(* Logix 5000 project; controller SigmaAldrich vendor 1 type 14 code 77 rev 15.4; software revision 15.02 *)

TASK MainTask (continuous, watchdog 500 ms) : MainProgram

MODULES
   Controller : vendor 1 type 14 code 77 (CompactLogixL32EController 0, rev 15.4)
      LocalENB : 1769-L32E Ethernet Port (CompactLogixL32Ethernet 1, rev 15.3)
      Local : CompactBus (CompactVirtualAdapter 3, rev 15.3, Input RPI 2 ms)
          : vendor 1 type 7 code 69 (Compact 12, rev 3.1, Input RPI 2 ms)
          : vendor 1 type 7 code 69 (Compact 9, rev 3.1, Input RPI 2 ms)
          : vendor 1 type 7 code 69 (Compact 7, rev 3.1, Input RPI 2 ms)
          : vendor 1 type 7 code 69 (Compact 10, rev 3.1, Input RPI 2 ms)
          : vendor 1 type 7 code 69 (Compact 11, rev 3.1, Input RPI 2 ms)
          : vendor 1 type 7 code 69 (Compact 8, rev 3.1, Input RPI 2 ms)
          : 1769-OW16 (Compact 1, rev 1.1, Output RPI 2 ms)
          : 1769-OW16 (Compact 6, rev 1.1, Output RPI 2 ms)
          : 1769-OW16 (Compact 3, rev 1.1, Output RPI 2 ms)
          : 1769-OW16 (Compact 4, rev 1.1, Output RPI 2 ms)
          : 1769-OW16 (Compact 2, rev 1.1, Output RPI 2 ms)
          : 1769-OW16 (Compact 5, rev 1.1, Output RPI 2 ms)
END_MODULES

VAR_GLOBAL   (* controller tags *)
   Airlock_N1002_03_04_E_Stop_OSR : BOOL;
   Airlock_N1002_03_04_Violation_MDI_Bit : BOOL := 1;
   Airlock_N1002_03_04_Violation_MDI_OSR : BOOL := 1;
   Airlock_N1005_E_Stop_OSR : BOOL;
   Airlock_N1005_Violation_MDI_Bit : BOOL;
   Airlock_N1005_Violation_MDI_OSR : BOOL;
   Airlock_N1006_E_Stop_OSR : BOOL;
   Airlock_N1006_Violation_MDI_Bit : BOOL;
   Airlock_N1006_Violation_MDI_OSR : BOOL;
   Airlock_N1008_E_Stop_OSR : BOOL;
   Airlock_N1008_Violation_MDI_Bit : BOOL;
   Airlock_N1008_Violation_MDI_OSR : BOOL;
   Airlock_N1009_E_Stop_OSR : BOOL;
   Airlock_N1009_Violation_MDI_Bit : BOOL;
   Airlock_N1009_Violation_MDI_OSR : BOOL;
   Airlock_N1011_E_Stop_OSR : BOOL;
   Airlock_N1011_Violation_MDI_Bit : BOOL := 1;
   Airlock_N1011_Violation_MDI_OSR : BOOL := 1;
   Airlock_N1012_E_Stop_OSR : BOOL;
   Airlock_N1012_Violation_MDI_Bit : BOOL := 1;
   Airlock_N1012_Violation_MDI_OSR : BOOL := 1;
   Airlock_N1021_E_Stop_OSR : BOOL;
   Airlock_N1021_Violation_MDI_Bit : BOOL;
   Airlock_N1021_Violation_MDI_OSR : BOOL;
   Airlock_N1043_E_Stop_OSR : BOOL;
   Airlock_N1043_Violation_MDI_Bit : BOOL := 1;
   Airlock_N1043_Violation_MDI_OSR : BOOL := 1;
   Airlock_N1044_E_Stop_OSR : BOOL;
   Airlock_N1044_Violation_MDI_Bit : BOOL;
   Airlock_N1044_Violation_MDI_OSR : BOOL;
   Airlock_N1051_54_55_E_Stop_OSR : BOOL;
   Airlock_N1051_54_55_Violation_MDI_Bit : BOOL := 1;
   Airlock_N1051_54_55_Violation_MDI_OSR : BOOL;
   Airlock_N1052_E_Stop_OSR : BOOL;
   Airlock_N1052_Violation_MDI_Bit : BOOL;
   Airlock_N1052_Violation_MDI_OSR : BOOL;
   Airlock_N1065_E_Stop_OSR : BOOL;
   Airlock_N1065_Violation_MDI_Bit : BOOL;
   Airlock_N1065_Violation_MDI_OSR : BOOL;
   Airlock_N1066_E_Stop_OSR : BOOL;
   Airlock_N1066_Violation_MDI_Bit : BOOL := 1;
   Airlock_N1066_Violation_MDI_OSR : BOOL := 1;
   Airlock_N1068_E_Stop_OSR : BOOL;
   Airlock_N1068_Violation_MDI_Bit : BOOL;
   Airlock_N1068_Violation_MDI_OSR : BOOL;
   Annuciator_Bit_Airlock_N1002_03_04 : BOOL := 1;
   Annuciator_Bit_Airlock_N1005 : BOOL;
   Annuciator_Bit_Airlock_N1006 : BOOL;
   Annuciator_Bit_Airlock_N1008 : BOOL;
   Annuciator_Bit_Airlock_N1009 : BOOL;
   Annuciator_Bit_Airlock_N1011 : BOOL := 1;
   Annuciator_Bit_Airlock_N1012 : BOOL := 1;
   Annuciator_Bit_Airlock_N1021 : BOOL;
   Annuciator_Bit_Airlock_N1043 : BOOL := 1;
   Annuciator_Bit_Airlock_N1044 : BOOL;
   Annuciator_Bit_Airlock_N1051_54_55 : BOOL := 1;
   Annuciator_Bit_Airlock_N1052 : BOOL;
   Annuciator_Bit_Airlock_N1065 : BOOL;
   Annuciator_Bit_Airlock_N1066 : BOOL := 1;
   Annuciator_Bit_Airlock_N1068 : BOOL;
   Door_N1002A_Timer : TIMER := (PRE := 30000);
   Door_N1002B_Timer : TIMER := (PRE := 30000);
   Door_N1002C_Timer : TIMER := (PRE := 30000);
   Door_N1003A_Timer : TIMER := (PRE := 30000);
   Door_N1003C_Timer : TIMER := (PRE := 30000, ACC := 30000, EN := 1, DN := 1);
   Door_N1004A_Timer : TIMER := (PRE := 30000);
   Door_N1004B_Timer : TIMER := (PRE := 30000);
   Door_N1005A_Timer : TIMER := (PRE := 30000);
   Door_N1005B_Timer : TIMER := (PRE := 30000);
   Door_N1006A_Timer : TIMER := (PRE := 30000);
   Door_N1006B_Timer : TIMER := (PRE := 30000);
   Door_N1008A_Timer : TIMER := (PRE := 30000);
   Door_N1008B_Timer : TIMER := (PRE := 30000);
   Door_N1009A_Timer : TIMER := (PRE := 30000);
   Door_N1009B_Timer : TIMER := (PRE := 30000);
   Door_N1011A_Timer : TIMER := (PRE := 30000, ACC := 30000, EN := 1, DN := 1);
   Door_N1011B_Timer : TIMER := (PRE := 30000, ACC := 30000, EN := 1, DN := 1);
   Door_N1012_Timer : TIMER := (PRE := 30000, ACC := 30000, EN := 1, DN := 1);
   Door_N1021A_Timer : TIMER := (PRE := 30000);
   Door_N1021B_Timer : TIMER := (PRE := 30000);
   Door_N1021C_Timer : TIMER := (PRE := 30000);
   Door_N1043A_Timer : TIMER := (PRE := 30000, ACC := 30000, EN := 1, DN := 1);
   Door_N1043B_Timer : TIMER := (PRE := 30000);
   Door_N1044A_Timer : TIMER := (PRE := 30000);
   Door_N1044B_Timer : TIMER := (PRE := 30000);
   Door_N1044C_Timer : TIMER := (PRE := 30000);
   Door_N1051A_Timer : TIMER := (PRE := 30000, ACC := 30000, EN := 1, DN := 1);
   Door_N1051B_Timer : TIMER := (PRE := 30000, ACC := 30000, EN := 1, DN := 1);
   Door_N1052A_Timer : TIMER := (PRE := 30000);
   Door_N1052B_Timer : TIMER := (PRE := 30000);
   Door_N1053_Timer : TIMER := (PRE := 30000, ACC := 30000, EN := 1, DN := 1);
   Door_N1054A_Timer : TIMER := (PRE := 30000, ACC := 30000, EN := 1, DN := 1);
   Door_N1054B_Timer : TIMER := (PRE := 30000, ACC := 30000, EN := 1, DN := 1);
   Door_N1054C_Timer : TIMER := (PRE := 30000, ACC := 30000, EN := 1, DN := 1);
   Door_N1055_Timer : TIMER := (PRE := 30000, ACC := 30000, EN := 1, DN := 1);
   Door_N1058B_Timer : TIMER := (PRE := 30000);
   Door_N1065A_Timer : TIMER := (PRE := 30000);
   Door_N1065B_Timer : TIMER := (PRE := 30000);
   Door_N1066A_Timer : TIMER := (PRE := 30000, ACC := 30000, EN := 1, DN := 1);
   Door_N1066B_Timer : TIMER := (PRE := 30000, ACC := 30000, EN := 1, DN := 1);
   Door_N1068A_Timer : TIMER := (PRE := 30000);
   Door_N1068B_Timer : TIMER := (PRE := 30000);
   MDI_Violation_N1002_03_04_Bit : BOOL := 1;
   MDI_Violation_N1005_Bit : BOOL;
   MDI_Violation_N1006_Bit : BOOL;
   MDI_Violation_N1008_Bit : BOOL;
   MDI_Violation_N1009_Bit : BOOL;
   MDI_Violation_N1011_Bit : BOOL := 1;
   MDI_Violation_N1012_Bit : BOOL := 1;
   MDI_Violation_N1021_Bit : BOOL;
   MDI_Violation_N1043_Bit : BOOL := 1;
   MDI_Violation_N1044_Bit : BOOL;
   MDI_Violation_N1051_54_55_Bit : BOOL := 1;
   MDI_Violation_N1052_Bit : BOOL;
   MDI_Violation_N1065_Bit : BOOL;
   MDI_Violation_N1066_Bit : BOOL := 1;
   MDI_Violation_N1068_Bit : BOOL;
   N1002_03_04_Airlock_Latch : BOOL := 1;
   N1002_03_04_Emergency_Release_Latch : BOOL := 1;
   N1005_Airlock_Latch : BOOL;
   N1005_Emergency_Release_Latch : BOOL;
   N1006_Airlock_Latch : BOOL;
   N1006_Emergency_Release_Latch : BOOL;
   N1008_Airlock_Latch : BOOL;
   N1008_Emergency_Release_Latch : BOOL;
   N1009_Airlock_Latch : BOOL;
   N1009_Emergency_Release_Latch : BOOL;
   N1011_Airlock_Latch : BOOL := 1;
   N1011_Emergency_Release_Latch : BOOL;
   N1012_Airlock_Latch : BOOL := 1;
   N1012_Emergency_Release_Latch : BOOL;
   N1021_Airlock_Latch : BOOL;
   N1021_Emergency_Release_Latch : BOOL;
   N1021C_Door_Latch_Bit : BOOL;
   N1043_Airlock_Latch : BOOL;
   N1043_Emergency_Release_Latch : BOOL;
   N1044_Airlock_Latch : BOOL;
   N1044_Emergency_Release_Latch : BOOL;
   N1044A_Door_Latch_Bit : BOOL;
   N1051_54_55_Airlock_Latch : BOOL := 1;
   N1051_54_55_Emergency_Release_Latch : BOOL;
   N1052_Airlock_Latch : BOOL;
   N1052_Emergency_Release_Latch : BOOL;
   N1052A_Door_Latch_Bit : BOOL;
   N1065_Airlock_Latch : BOOL;
   N1065_Emergency_Release_Latch : BOOL;
   N1066_Airlock_Latch : BOOL := 1;
   N1066_Emergency_Release_Latch : BOOL;
   N1068_Airlock_Latch : BOOL;
   N1068_Emergency_Release_Latch : BOOL;
   N1068B_Door_Latch_Bit : BOOL;
END_VAR

PROGRAM MainProgram   (* main routine MainRoutine *)
VAR
   Airlock_N1009_Delay_Tmr : TIMER := (PRE := 2000);
   Airlock_N1009_MDI_Delay_Tmr : TIMER := (PRE := 2000, ACC := 2001, EN := 1, DN := 1);
END_VAR

ROUTINE DI01_N1051_N1054_N0155   (* ladder *)
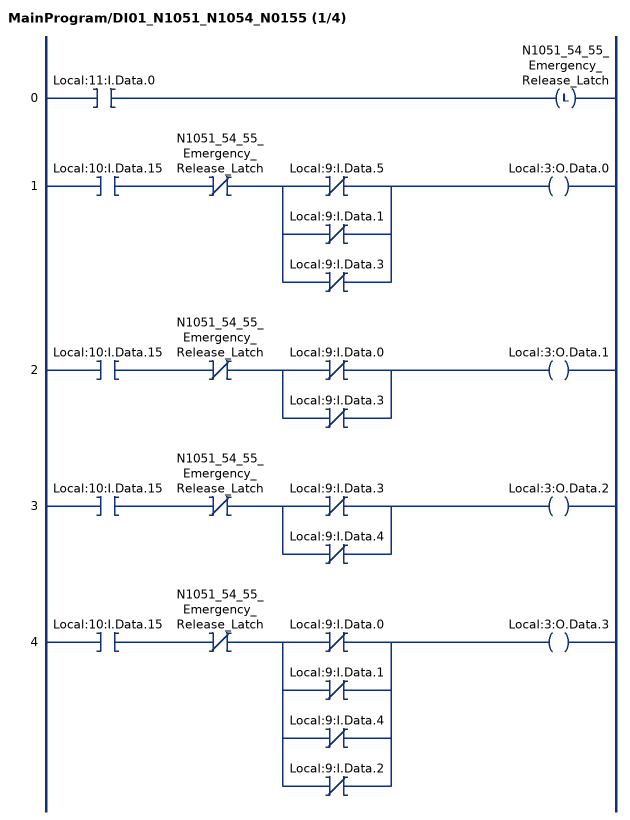
   0: XIC(Local:11:I.Data.0)OTL(N1051_54_55_Emergency_Release_Latch);
   1: XIC(Local:10:I.Data.15)XIO(N1051_54_55_Emergency_Release_Latch)[XIO(Local:9:I.Data.5) ,XIO(Local:9:I.Data.1) ,XIO(Local:9:I.Data.3) ]OTE(Local:3:O.Data.0);
   2: XIC(Local:10:I.Data.15)XIO(N1051_54_55_Emergency_Release_Latch)[XIO(Local:9:I.Data.0) ,XIO(Local:9:I.Data.3) ]OTE(Local:3:O.Data.1);
   3: XIC(Local:10:I.Data.15)XIO(N1051_54_55_Emergency_Release_Latch)[XIO(Local:9:I.Data.3) ,XIO(Local:9:I.Data.4) ]OTE(Local:3:O.Data.2);
   4: XIC(Local:10:I.Data.15)XIO(N1051_54_55_Emergency_Release_Latch)[XIO(Local:9:I.Data.0) ,XIO(Local:9:I.Data.1) ,XIO(Local:9:I.Data.4) ,XIO(Local:9:I.Data.2) ]OTE(Local:3:O.Data.3);
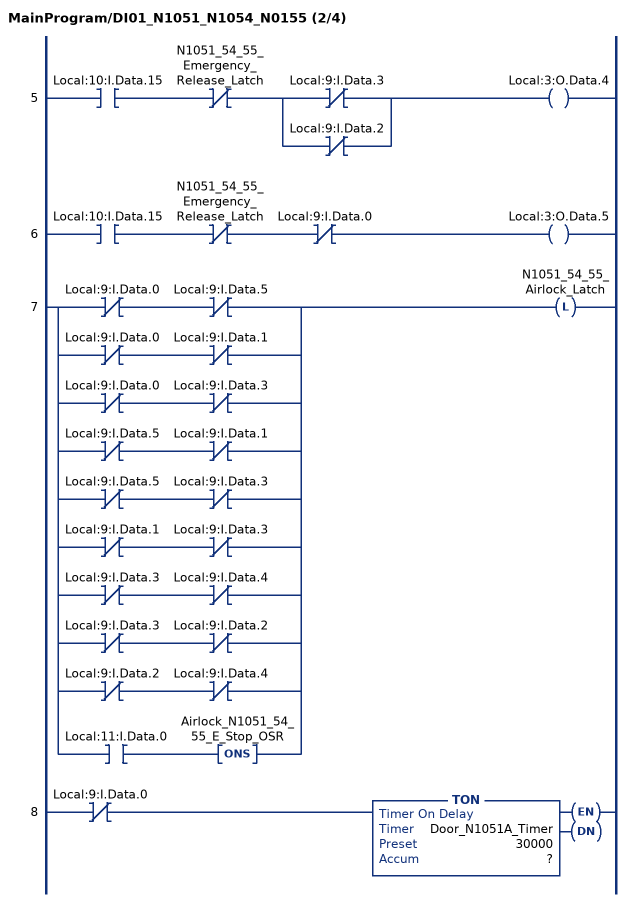
   5: XIC(Local:10:I.Data.15)XIO(N1051_54_55_Emergency_Release_Latch)[XIO(Local:9:I.Data.3) ,XIO(Local:9:I.Data.2) ]OTE(Local:3:O.Data.4);
   6: XIC(Local:10:I.Data.15)XIO(N1051_54_55_Emergency_Release_Latch)XIO(Local:9:I.Data.0)OTE(Local:3:O.Data.5);
   7: [XIO(Local:9:I.Data.0) XIO(Local:9:I.Data.5) ,XIO(Local:9:I.Data.0) XIO(Local:9:I.Data.1) ,XIO(Local:9:I.Data.0) XIO(Local:9:I.Data.3) ,XIO(Local:9:I.Data.5) XIO(Local:9:I.Data.1) ,XIO(Local:9:I.Data.5) XIO(Local:9:I.Data.3) ,XIO(Local:9:I.Data.1) XIO(Local:9:I.Data.3) ,XIO(Local:9:I.Data.3) XIO(Local:9:I.Data.4) ,XIO(Local:9:I.Data.3) XIO(Local:9:I.Data.2) ,XIO(Local:9:I.Data.2) XIO(Local:9:I.Data.4) ,XIC(Local:11:I.Data.0) ONS(Airlock_N1051_54_55_E_Stop_OSR) ]OTL(N1051_54_55_Airlock_Latch);
   8: XIO(Local:9:I.Data.0)TON(Door_N1051A_Timer,?,?);
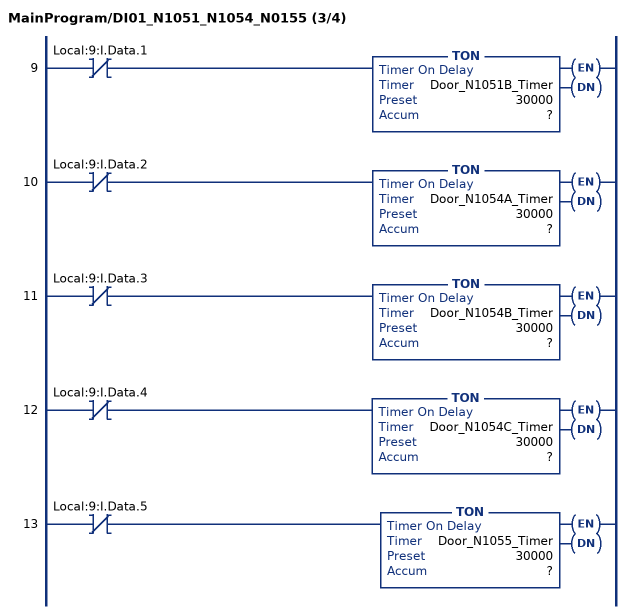
   9: XIO(Local:9:I.Data.1)TON(Door_N1051B_Timer,?,?);
   10: XIO(Local:9:I.Data.2)TON(Door_N1054A_Timer,?,?);
   11: XIO(Local:9:I.Data.3)TON(Door_N1054B_Timer,?,?);
   12: XIO(Local:9:I.Data.4)TON(Door_N1054C_Timer,?,?);
   13: XIO(Local:9:I.Data.5)TON(Door_N1055_Timer,?,?);
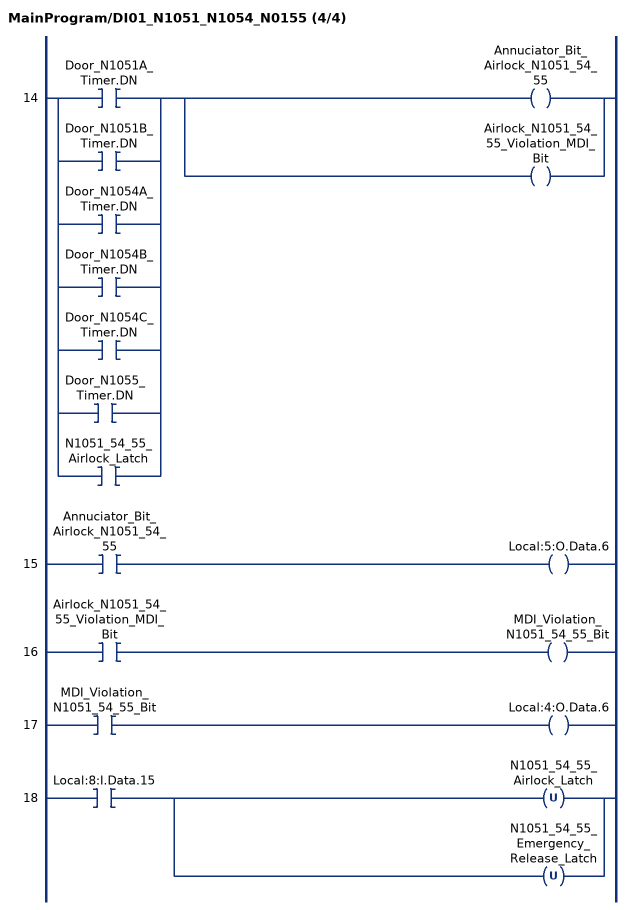
   14: [XIC(Door_N1051A_Timer.DN) ,XIC(Door_N1051B_Timer.DN) ,XIC(Door_N1054A_Timer.DN) ,XIC(Door_N1054B_Timer.DN) ,XIC(Door_N1054C_Timer.DN) ,XIC(Door_N1055_Timer.DN) ,XIC(N1051_54_55_Airlock_Latch) ][OTE(Annuciator_Bit_Airlock_N1051_54_55) ,OTE(Airlock_N1051_54_55_Violation_MDI_Bit) ];
   15: XIC(Annuciator_Bit_Airlock_N1051_54_55)OTE(Local:5:O.Data.6);
   16: XIC(Airlock_N1051_54_55_Violation_MDI_Bit)OTE(MDI_Violation_N1051_54_55_Bit);
   17: XIC(MDI_Violation_N1051_54_55_Bit)OTE(Local:4:O.Data.6);
   18: XIC(Local:8:I.Data.15)[OTU(N1051_54_55_Airlock_Latch) ,OTU(N1051_54_55_Emergency_Release_Latch) ];
END_ROUTINE

ROUTINE DI02_N1002_N1003_N1004   (* ladder *)
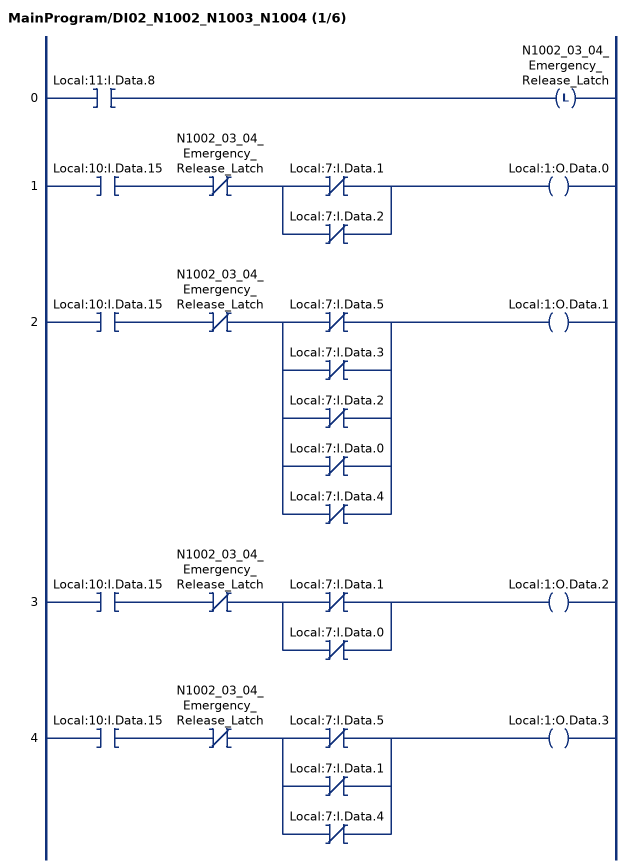
   0: XIC(Local:11:I.Data.8)OTL(N1002_03_04_Emergency_Release_Latch);
   1: XIC(Local:10:I.Data.15)XIO(N1002_03_04_Emergency_Release_Latch)[XIO(Local:7:I.Data.1) ,XIO(Local:7:I.Data.2) ]OTE(Local:1:O.Data.0);
   2: XIC(Local:10:I.Data.15)XIO(N1002_03_04_Emergency_Release_Latch)[XIO(Local:7:I.Data.5) ,XIO(Local:7:I.Data.3) ,XIO(Local:7:I.Data.2) ,XIO(Local:7:I.Data.0) ,XIO(Local:7:I.Data.4) ]OTE(Local:1:O.Data.1);
   3: XIC(Local:10:I.Data.15)XIO(N1002_03_04_Emergency_Release_Latch)[XIO(Local:7:I.Data.1) ,XIO(Local:7:I.Data.0) ]OTE(Local:1:O.Data.2);
   4: XIC(Local:10:I.Data.15)XIO(N1002_03_04_Emergency_Release_Latch)[XIO(Local:7:I.Data.5) ,XIO(Local:7:I.Data.1) ,XIO(Local:7:I.Data.4) ]OTE(Local:1:O.Data.3);
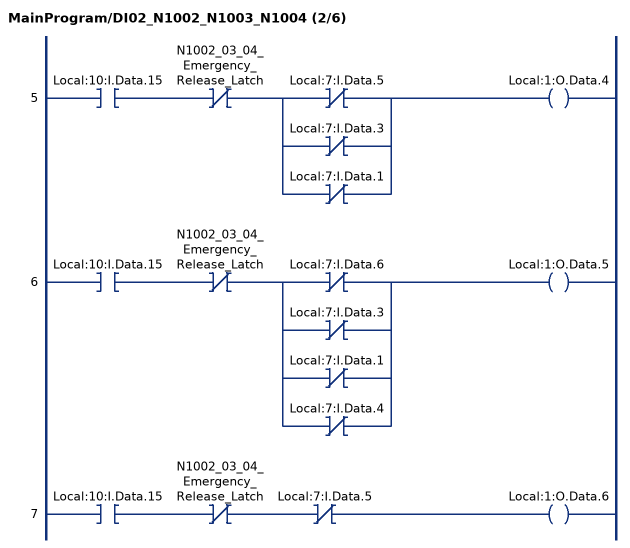
   5: XIC(Local:10:I.Data.15)XIO(N1002_03_04_Emergency_Release_Latch)[XIO(Local:7:I.Data.5) ,XIO(Local:7:I.Data.3) ,XIO(Local:7:I.Data.1) ]OTE(Local:1:O.Data.4);
   6: XIC(Local:10:I.Data.15)XIO(N1002_03_04_Emergency_Release_Latch)[XIO(Local:7:I.Data.6) ,XIO(Local:7:I.Data.3) ,XIO(Local:7:I.Data.1) ,XIO(Local:7:I.Data.4) ]OTE(Local:1:O.Data.5);
   7: XIC(Local:10:I.Data.15)XIO(N1002_03_04_Emergency_Release_Latch)XIO(Local:7:I.Data.5)OTE(Local:1:O.Data.6);
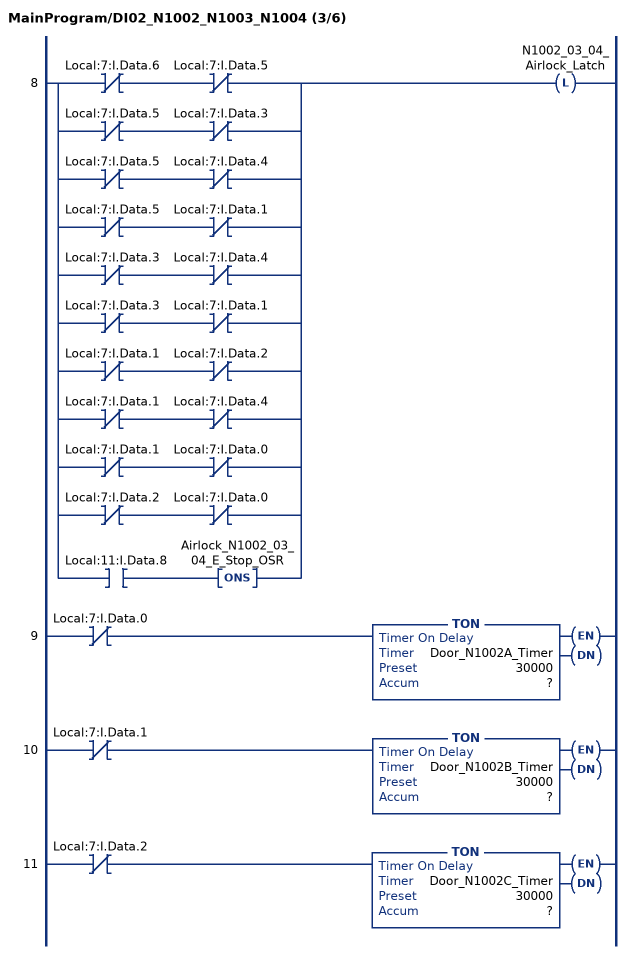
   8: [XIO(Local:7:I.Data.6) XIO(Local:7:I.Data.5) ,XIO(Local:7:I.Data.5) XIO(Local:7:I.Data.3) ,XIO(Local:7:I.Data.5) XIO(Local:7:I.Data.4) ,XIO(Local:7:I.Data.5) XIO(Local:7:I.Data.1) ,XIO(Local:7:I.Data.3) XIO(Local:7:I.Data.4) ,XIO(Local:7:I.Data.3) XIO(Local:7:I.Data.1) ,XIO(Local:7:I.Data.1) XIO(Local:7:I.Data.2) ,XIO(Local:7:I.Data.1) XIO(Local:7:I.Data.4) ,XIO(Local:7:I.Data.1) XIO(Local:7:I.Data.0) ,XIO(Local:7:I.Data.2) XIO(Local:7:I.Data.0) ,XIC(Local:11:I.Data.8) ONS(Airlock_N1002_03_04_E_Stop_OSR) ]OTL(N1002_03_04_Airlock_Latch);
   9: XIO(Local:7:I.Data.0)TON(Door_N1002A_Timer,?,?);
   10: XIO(Local:7:I.Data.1)TON(Door_N1002B_Timer,?,?);
   11: XIO(Local:7:I.Data.2)TON(Door_N1002C_Timer,?,?);
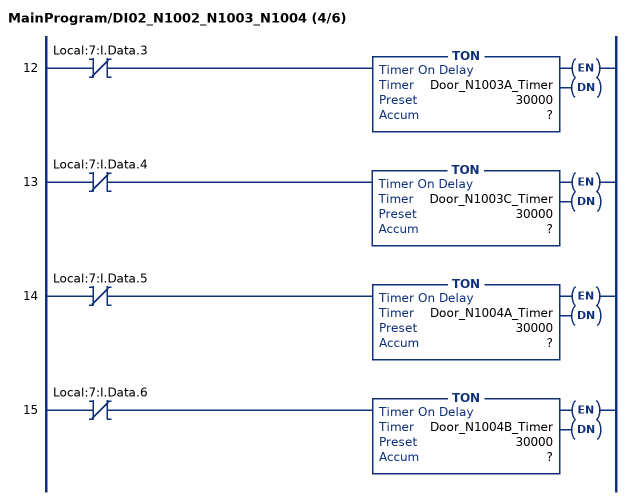
   12: XIO(Local:7:I.Data.3)TON(Door_N1003A_Timer,?,?);
   13: XIO(Local:7:I.Data.4)TON(Door_N1003C_Timer,?,?);
   14: XIO(Local:7:I.Data.5)TON(Door_N1004A_Timer,?,?);
   15: XIO(Local:7:I.Data.6)TON(Door_N1004B_Timer,?,?);
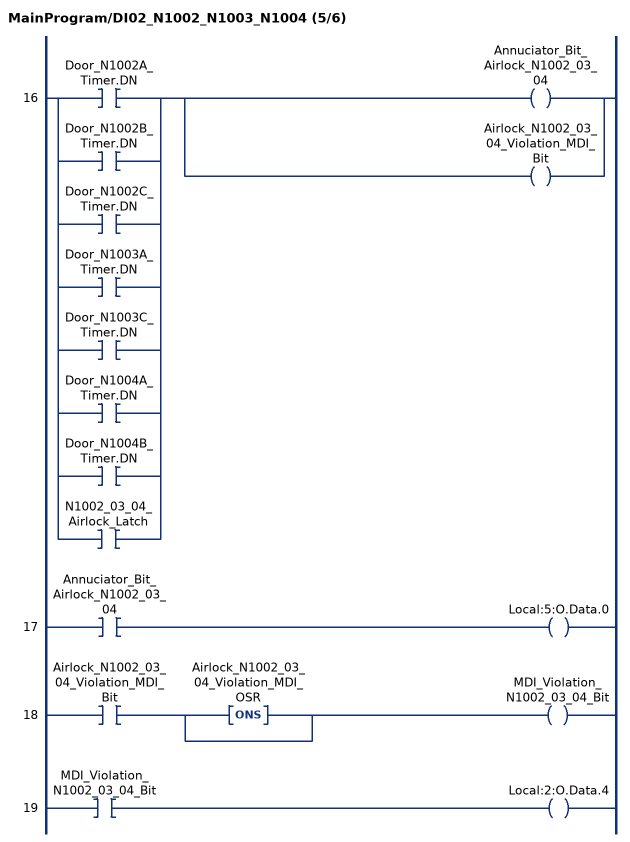
   16: [XIC(Door_N1002A_Timer.DN) ,XIC(Door_N1002B_Timer.DN) ,XIC(Door_N1002C_Timer.DN) ,XIC(Door_N1003A_Timer.DN) ,XIC(Door_N1003C_Timer.DN) ,XIC(Door_N1004A_Timer.DN) ,XIC(Door_N1004B_Timer.DN) ,XIC(N1002_03_04_Airlock_Latch) ][OTE(Annuciator_Bit_Airlock_N1002_03_04) ,OTE(Airlock_N1002_03_04_Violation_MDI_Bit) ];
   17: XIC(Annuciator_Bit_Airlock_N1002_03_04)OTE(Local:5:O.Data.0);
   18: XIC(Airlock_N1002_03_04_Violation_MDI_Bit)[ONS(Airlock_N1002_03_04_Violation_MDI_OSR) ,]OTE(MDI_Violation_N1002_03_04_Bit);
   19: XIC(MDI_Violation_N1002_03_04_Bit)OTE(Local:2:O.Data.4);
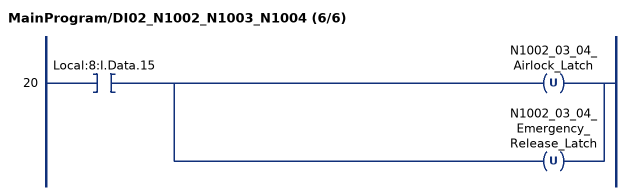
   20: XIC(Local:8:I.Data.15)[OTU(N1002_03_04_Airlock_Latch) ,OTU(N1002_03_04_Emergency_Release_Latch) ];
END_ROUTINE

ROUTINE DI03_N1021   (* ladder *)
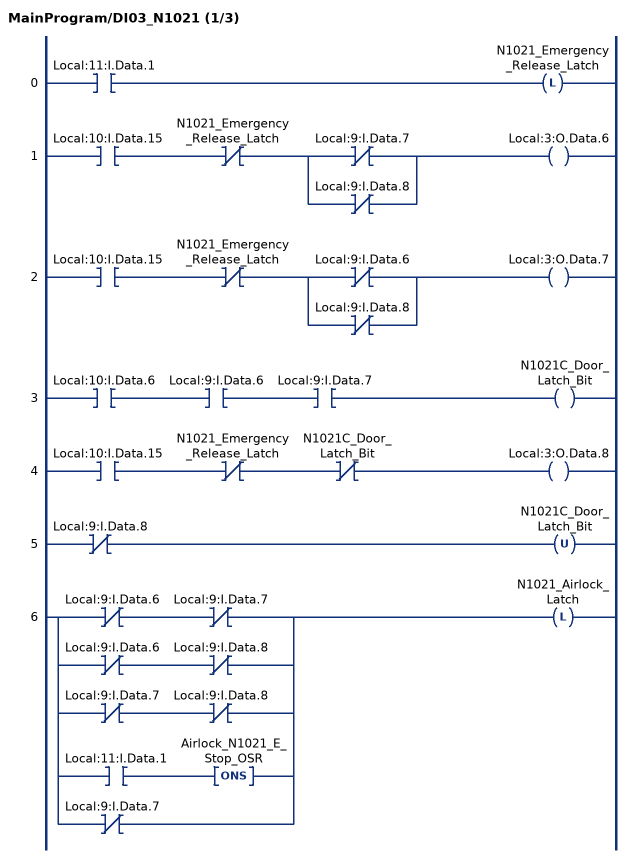
   0: XIC(Local:11:I.Data.1)OTL(N1021_Emergency_Release_Latch);
   1: XIC(Local:10:I.Data.15)XIO(N1021_Emergency_Release_Latch)[XIO(Local:9:I.Data.7) ,XIO(Local:9:I.Data.8) ]OTE(Local:3:O.Data.6);
   2: XIC(Local:10:I.Data.15)XIO(N1021_Emergency_Release_Latch)[XIO(Local:9:I.Data.6) ,XIO(Local:9:I.Data.8) ]OTE(Local:3:O.Data.7);
   3: XIC(Local:10:I.Data.6)XIC(Local:9:I.Data.6)XIC(Local:9:I.Data.7)OTE(N1021C_Door_Latch_Bit);
   4: XIC(Local:10:I.Data.15)XIO(N1021_Emergency_Release_Latch)XIO(N1021C_Door_Latch_Bit)OTE(Local:3:O.Data.8);
   5: XIO(Local:9:I.Data.8)OTU(N1021C_Door_Latch_Bit);
   6: [XIO(Local:9:I.Data.6) XIO(Local:9:I.Data.7) ,XIO(Local:9:I.Data.6) XIO(Local:9:I.Data.8) ,XIO(Local:9:I.Data.7) XIO(Local:9:I.Data.8) ,XIC(Local:11:I.Data.1) ONS(Airlock_N1021_E_Stop_OSR) ,XIO(Local:9:I.Data.7) ]OTL(N1021_Airlock_Latch);
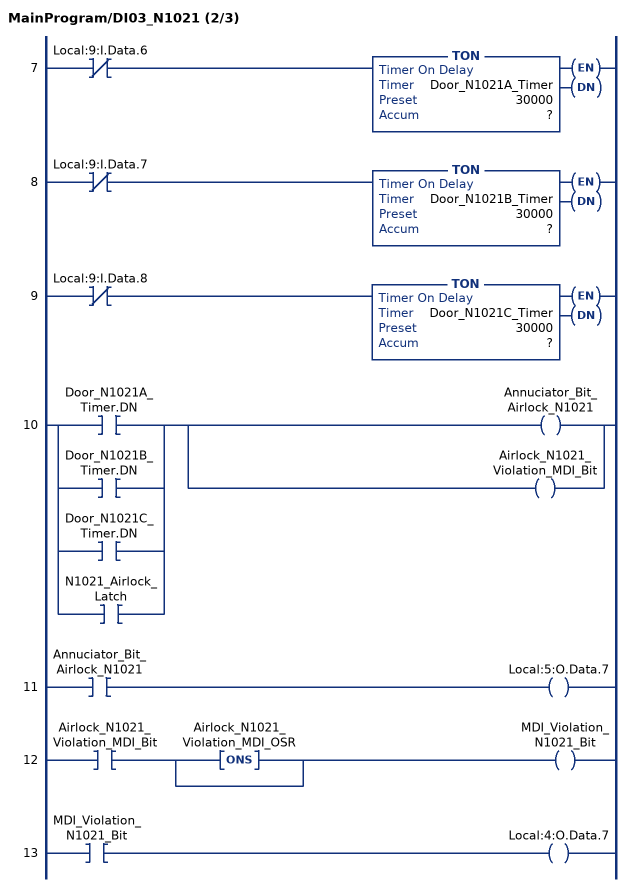
   7: XIO(Local:9:I.Data.6)TON(Door_N1021A_Timer,?,?);
   8: XIO(Local:9:I.Data.7)TON(Door_N1021B_Timer,?,?);
   9: XIO(Local:9:I.Data.8)TON(Door_N1021C_Timer,?,?);
   10: [XIC(Door_N1021A_Timer.DN) ,XIC(Door_N1021B_Timer.DN) ,XIC(Door_N1021C_Timer.DN) ,XIC(N1021_Airlock_Latch) ][OTE(Annuciator_Bit_Airlock_N1021) ,OTE(Airlock_N1021_Violation_MDI_Bit) ];
   11: XIC(Annuciator_Bit_Airlock_N1021)OTE(Local:5:O.Data.7);
   12: XIC(Airlock_N1021_Violation_MDI_Bit)[ONS(Airlock_N1021_Violation_MDI_OSR) ,]OTE(MDI_Violation_N1021_Bit);
   13: XIC(MDI_Violation_N1021_Bit)OTE(Local:4:O.Data.7);
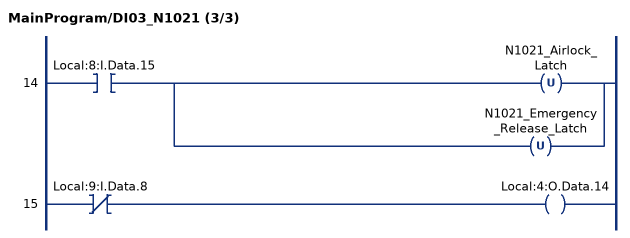
   14: XIC(Local:8:I.Data.15)[OTU(N1021_Airlock_Latch) ,OTU(N1021_Emergency_Release_Latch) ];
   15: XIO(Local:9:I.Data.8)OTE(Local:4:O.Data.14);
END_ROUTINE

ROUTINE DI04_N1005   (* ladder *)
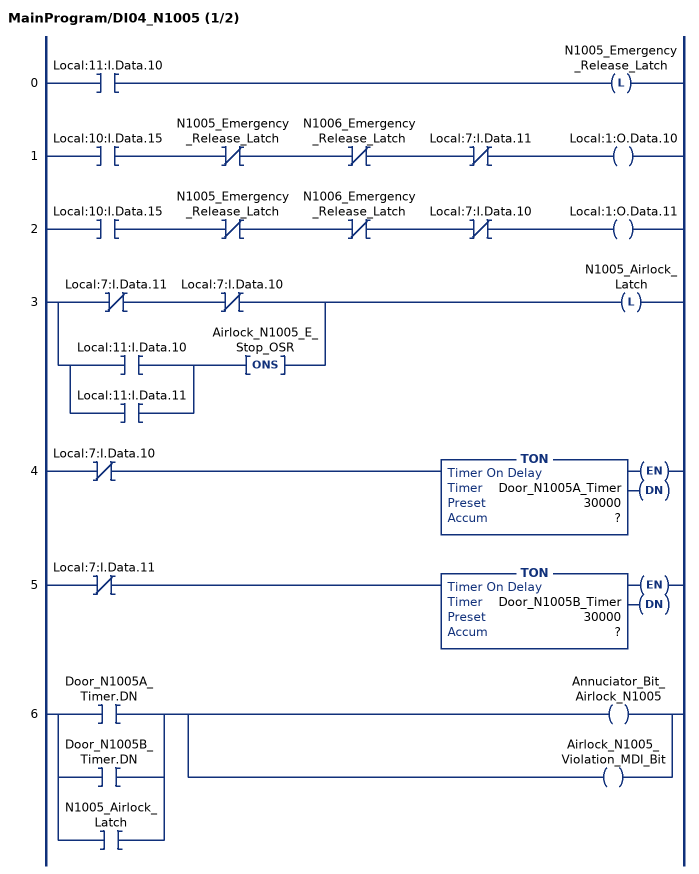
   0: XIC(Local:11:I.Data.10)OTL(N1005_Emergency_Release_Latch);
   1: XIC(Local:10:I.Data.15)XIO(N1005_Emergency_Release_Latch)XIO(N1006_Emergency_Release_Latch)XIO(Local:7:I.Data.11)OTE(Local:1:O.Data.10);
   2: XIC(Local:10:I.Data.15)XIO(N1005_Emergency_Release_Latch)XIO(N1006_Emergency_Release_Latch)XIO(Local:7:I.Data.10)OTE(Local:1:O.Data.11);
   3: [XIO(Local:7:I.Data.11) XIO(Local:7:I.Data.10) ,[XIC(Local:11:I.Data.10) ,XIC(Local:11:I.Data.11) ] ONS(Airlock_N1005_E_Stop_OSR) ]OTL(N1005_Airlock_Latch);
   4: XIO(Local:7:I.Data.10)TON(Door_N1005A_Timer,?,?);
   5: XIO(Local:7:I.Data.11)TON(Door_N1005B_Timer,?,?);
   6: [XIC(Door_N1005A_Timer.DN) ,XIC(Door_N1005B_Timer.DN) ,XIC(N1005_Airlock_Latch) ][OTE(Annuciator_Bit_Airlock_N1005) ,OTE(Airlock_N1005_Violation_MDI_Bit) ];
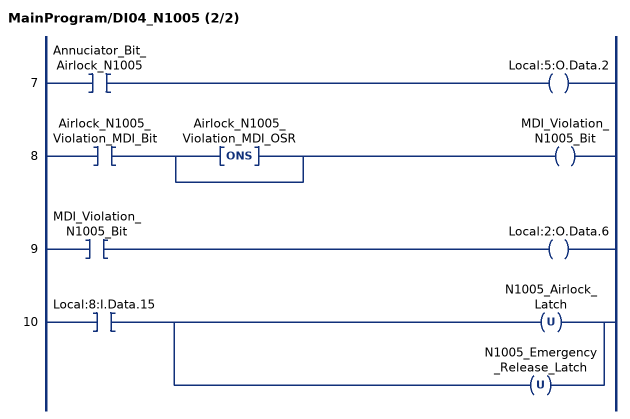
   7: XIC(Annuciator_Bit_Airlock_N1005)OTE(Local:5:O.Data.2);
   8: XIC(Airlock_N1005_Violation_MDI_Bit)[ONS(Airlock_N1005_Violation_MDI_OSR) ,]OTE(MDI_Violation_N1005_Bit);
   9: XIC(MDI_Violation_N1005_Bit)OTE(Local:2:O.Data.6);
   10: XIC(Local:8:I.Data.15)[OTU(N1005_Airlock_Latch) ,OTU(N1005_Emergency_Release_Latch) ];
END_ROUTINE

ROUTINE DI05_N1006   (* ladder *)
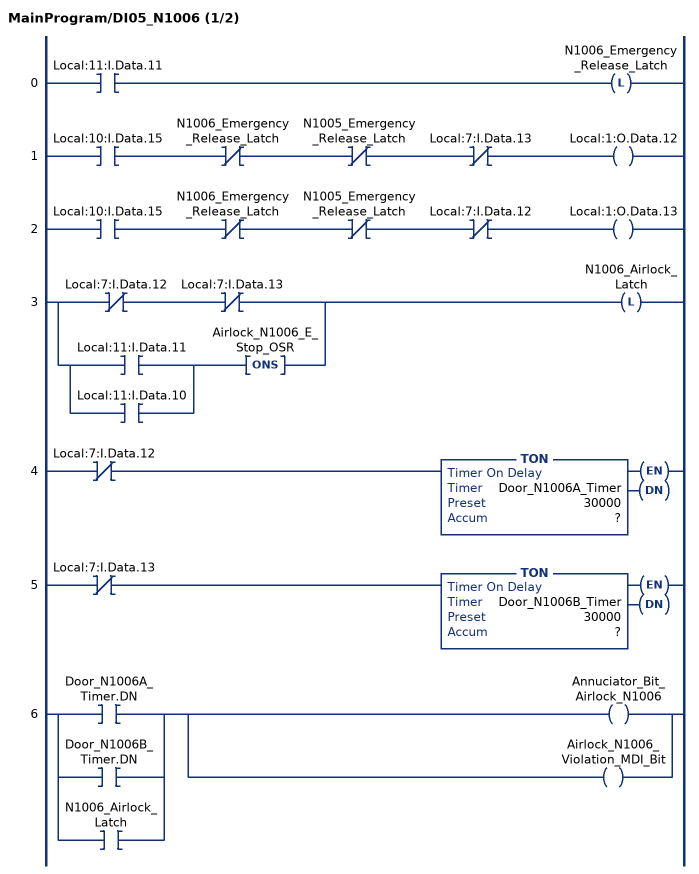
   0: XIC(Local:11:I.Data.11)OTL(N1006_Emergency_Release_Latch);
   1: XIC(Local:10:I.Data.15)XIO(N1006_Emergency_Release_Latch)XIO(N1005_Emergency_Release_Latch)XIO(Local:7:I.Data.13)OTE(Local:1:O.Data.12);
   2: XIC(Local:10:I.Data.15)XIO(N1006_Emergency_Release_Latch)XIO(N1005_Emergency_Release_Latch)XIO(Local:7:I.Data.12)OTE(Local:1:O.Data.13);
   3: [XIO(Local:7:I.Data.12) XIO(Local:7:I.Data.13) ,[XIC(Local:11:I.Data.11) ,XIC(Local:11:I.Data.10) ] ONS(Airlock_N1006_E_Stop_OSR) ]OTL(N1006_Airlock_Latch);
   4: XIO(Local:7:I.Data.12)TON(Door_N1006A_Timer,?,?);
   5: XIO(Local:7:I.Data.13)TON(Door_N1006B_Timer,?,?);
   6: [XIC(Door_N1006A_Timer.DN) ,XIC(Door_N1006B_Timer.DN) ,XIC(N1006_Airlock_Latch) ][OTE(Annuciator_Bit_Airlock_N1006) ,OTE(Airlock_N1006_Violation_MDI_Bit) ];
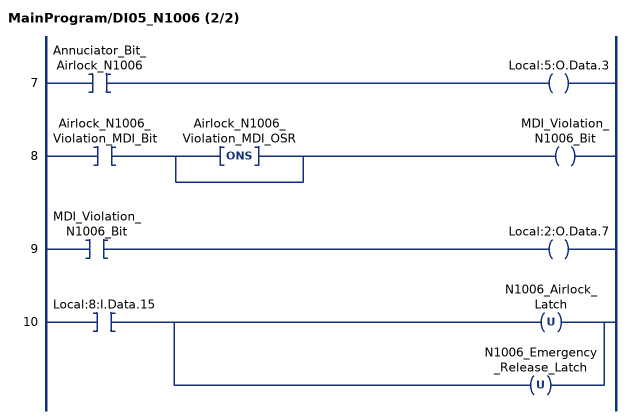
   7: XIC(Annuciator_Bit_Airlock_N1006)OTE(Local:5:O.Data.3);
   8: XIC(Airlock_N1006_Violation_MDI_Bit)[ONS(Airlock_N1006_Violation_MDI_OSR) ,]OTE(MDI_Violation_N1006_Bit);
   9: XIC(MDI_Violation_N1006_Bit)OTE(Local:2:O.Data.7);
   10: XIC(Local:8:I.Data.15)[OTU(N1006_Airlock_Latch) ,OTU(N1006_Emergency_Release_Latch) ];
END_ROUTINE

ROUTINE DI06_N1008   (* ladder *)
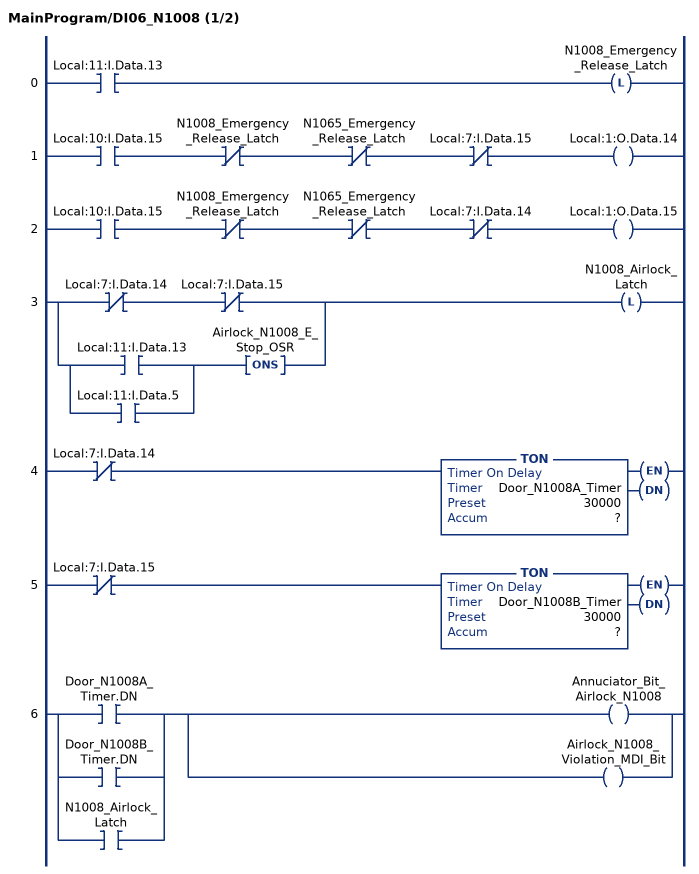
   0: XIC(Local:11:I.Data.13)OTL(N1008_Emergency_Release_Latch);
   1: XIC(Local:10:I.Data.15)XIO(N1008_Emergency_Release_Latch)XIO(N1065_Emergency_Release_Latch)XIO(Local:7:I.Data.15)OTE(Local:1:O.Data.14);
   2: XIC(Local:10:I.Data.15)XIO(N1008_Emergency_Release_Latch)XIO(N1065_Emergency_Release_Latch)XIO(Local:7:I.Data.14)OTE(Local:1:O.Data.15);
   3: [XIO(Local:7:I.Data.14) XIO(Local:7:I.Data.15) ,[XIC(Local:11:I.Data.13) ,XIC(Local:11:I.Data.5) ] ONS(Airlock_N1008_E_Stop_OSR) ]OTL(N1008_Airlock_Latch);
   4: XIO(Local:7:I.Data.14)TON(Door_N1008A_Timer,?,?);
   5: XIO(Local:7:I.Data.15)TON(Door_N1008B_Timer,?,?);
   6: [XIC(Door_N1008A_Timer.DN) ,XIC(Door_N1008B_Timer.DN) ,XIC(N1008_Airlock_Latch) ][OTE(Annuciator_Bit_Airlock_N1008) ,OTE(Airlock_N1008_Violation_MDI_Bit) ];
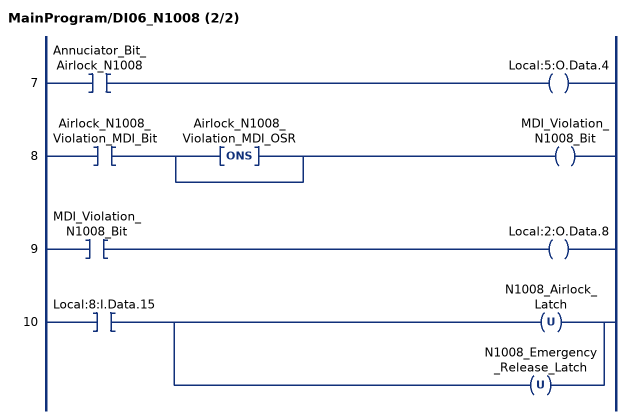
   7: XIC(Annuciator_Bit_Airlock_N1008)OTE(Local:5:O.Data.4);
   8: XIC(Airlock_N1008_Violation_MDI_Bit)[ONS(Airlock_N1008_Violation_MDI_OSR) ,]OTE(MDI_Violation_N1008_Bit);
   9: XIC(MDI_Violation_N1008_Bit)OTE(Local:2:O.Data.8);
   10: XIC(Local:8:I.Data.15)[OTU(N1008_Airlock_Latch) ,OTU(N1008_Emergency_Release_Latch) ];
END_ROUTINE
